Fanuc KAREL source: kb00003.compact.KL

PROGRAM KB00003
%STACKSIZE=65535
%PRIORITY=65535
%NOLOCKGROUP
VAR
P1 : REAL
RESULT : REAL
BEGIN
P1=1.0
RESULT=ACOS(P1)
END KB00003
